(* IEC 61131-3 sources: rusty/tests/lit/single/arithmetic, 10 files *)

(* ---- addition.st ---- *)
// RUN: %COMPILE %s && %RUN | %CHECK %s
// CHECK: 10
FUNCTION main
    VAR
        x : DINT;
        y : DINT;
    END_VAR

    x := 5;
    y := 5;
    printf('%d$N', x + y);
END_FUNCTION

(* ---- integer_overflow.st ---- *)
// RUN: %COMPILE %s && %RUN | %CHECK %s
FUNCTION main
    VAR
        var_sint    : SINT;
        var_int     : INT;
        var_dint    : DINT;
        var_lint    : LINT;

        var_usint   : USINT;
        var_uint    : UINT;
        var_udint   : UDINT;
        var_ulint   : ULINT;
    END_VAR

    // Set max values
    // 8-bit [(2^7)-1]/[(2^8)-1]
    var_sint := 127;                    // Min: -128
    var_usint := 255;                   // Min: 0

    // 16-bit [(2^15)-1]/[(2^16)-1]
    var_int := 32767;                   // Min: -32768
    var_uint := 65535;                  // Min: 0

    // 32-bit [(2^31)-1]/[(2^31)-1]
    var_dint := 2147483647;             // Min: -2147483648
    var_udint := 4294967295;            // Min: 0

    // 64-bit [(2^63)-1]/[(2^64)-1]
    var_lint := 9223372036854775807;    // Min: -9223372036854775808
    var_ulint := 18446744073709551615;  // Min: 0

    // Print and check values
    printf('%d$N', var_sint);       // CHECK: 127
    printf('%d$N', var_int);        // CHECK-NEXT: 32767
    printf('%d$N', var_dint);       // CHECK-NEXT: 2147483647
    printf('%lld$N', var_lint);     // CHECK-NEXT: 9223372036854775807

    printf('%u$N', var_usint);      // CHECK-NEXT: 255
    printf('%u$N', var_uint);       // CHECK-NEXT: 65535
    printf('%u$N', var_udint);      // CHECK-NEXT: 4294967295
    printf('%llu$N', var_ulint);    // CHECK-NEXT: 18446744073709551615

    // Print overflow values
    var_sint := var_sint + 1;
    var_int := var_int + 1;
    var_dint := var_dint + 1;
    var_lint := var_lint + 1;

    var_usint := var_usint + 1;
    var_uint := var_uint + 1;
    var_udint := var_udint + 1;
    var_ulint := var_ulint + 1;

    printf('%d$N', var_sint);       // CHECK: -128
    printf('%d$N', var_int);        // CHECK-NEXT: -32768
    printf('%d$N', var_dint);       // CHECK-NEXT: -2147483648
    printf('%lld$N', var_lint);     // CHECK-NEXT: -9223372036854775808

    printf('%u$N', var_usint);      // CHECK-NEXT: 0
    printf('%u$N', var_uint);       // CHECK-NEXT: 0
    printf('%u$N', var_udint);      // CHECK-NEXT: 0
    printf('%llu$N', var_ulint);    // CHECK-NEXT: 0

END_FUNCTION

(* ---- integer_overflow_with_real_cast.st ---- *)
// RUN: %COMPILE %s && %RUN | %CHECK %s
FUNCTION main
    VAR
        var_int     : INT;
    END_VAR

    printf('%d$N', var_int); // CHECK: 0

    // Cast the REAL value to INT
    var_int := REAL_TO_INT(70_000.4);

    printf('%d$N', var_int); // CHECK: 32767

END_FUNCTION

(* ---- replaced_expression_result_cast.st ---- *)
// RUN: %COMPILE %s && %RUN | %CHECK %s
// The result of a builtin or an operator the compiler carries out through a function call is
// converted to the type of the variable it is assigned to

FUNCTION main
    VAR
        t : TIME := T#10s;
        lt : LTIME := LTIME#10s;
        tod : TOD := TOD#23:59:50;
        n : DINT := 7;
        m : DINT := 3;
        i : INT;
        r : REAL := 2.5;
        x : LREAL;
    END_VAR

    x := t * 1.5;
    printf('%.1f$N', x);                                                            // CHECK: 15000.0
    r := t / 4.0;
    x := r;
    printf('%.1f$N', x);                                                            // CHECK: 2500.0
    x := lt + lt;
    printf('%.1f$N', x);                                                            // CHECK: 20000000000.0

    x := MUL(t, 1.5);
    printf('%.1f$N', x);                                                            // CHECK: 15000.0
    x := ADD(n, m);
    printf('%.1f$N', x);                                                            // CHECK: 10.0
    r := 2.5;
    n := ADD(n, r);
    printf('%d$N', n);                                                              // CHECK: 9
    i := SUB(t, T#4s);
    printf('%d$N', i);                                                              // CHECK: 6000

    tod := (tod + T#20s);
    printf('%s$N', REF(TOD_TO_STRING(tod)));                                        // CHECK: TOD#00:00:10

END_FUNCTION

(* ---- sqrt.st ---- *)
// RUN: %COMPILE %s && %RUN | %CHECK %s
// CHECK: 2
FUNCTION main
    VAR
        res : LREAL;
    END_VAR
    printf('%d$N', REAL_TO_DINT(SQRT(4.0)));
END_FUNCTION

(* ---- unsigned_division_by_literal.st ---- *)
// RUN: %COMPILE %s && %RUN | %CHECK %s
//
// A division of an unsigned operand of 32 or 64 bits by an integer literal is unsigned, like a
// division by a variable of the same type, also when the operand has the highest bit set.

FUNCTION main
    VAR
        udint_value : UDINT := 4_000_000_000;
        two : UDINT := 2;
        dword_value : DWORD := 16#FFFF_FFFF;
        ulint_value : ULINT := 18_446_744_073_709_551_615;
        lword_value : LWORD := 16#FFFF_FFFF_FFFF_FFFF;
    END_VAR
    printf('udint / two: %u$N', udint_value / two);
    printf('udint / 2: %u$N', udint_value / 2);
    printf('dword / 2: %u$N', dword_value / 2);
    printf('ulint / 2: %llu$N', ulint_value / 2);
    printf('lword / 2: %llu$N', lword_value / 2);
    // CHECK:      udint / two: 2000000000
    // CHECK-NEXT: udint / 2: 2000000000
    // CHECK-NEXT: dword / 2: 2147483647
    // CHECK-NEXT: ulint / 2: 9223372036854775807
    // CHECK-NEXT: lword / 2: 9223372036854775807
END_FUNCTION

(* ---- unsigned_division_by_negative_literal.st ---- *)
// RUN: %COMPILE %s && %RUN | %CHECK %s
//
// A negative integer literal does not fit into an unsigned type, so a division or MOD of a UDINT by
// it still runs in DINT and gives a signed result.

FUNCTION main
    VAR
        value : UDINT := 10;
    END_VAR
    printf('value / -2: %d$N', value / -2);
    printf('value MOD -3: %d$N', value MOD -3);
    // CHECK:      value / -2: -5
    // CHECK-NEXT: value MOD -3: 1
END_FUNCTION

(* ---- unsigned_literal_dividend.st ---- *)
// RUN: %COMPILE %s && %RUN | %CHECK %s
//
// An integer literal as the left operand of a division or MOD takes the type of an unsigned divisor of
// 32 bits, so a divisor with the highest bit set is not read as a negative number. As a DINT,
// 16#FFFF_FFFF would be -1, and the results would be -100 and 0.

FUNCTION main
    VAR
        divisor : UDINT := 16#FFFF_FFFF;
    END_VAR
    printf('100 / divisor: %u$N', 100 / divisor);
    printf('100 MOD divisor: %u$N', 100 MOD divisor);
    // CHECK:      100 / divisor: 0
    // CHECK-NEXT: 100 MOD divisor: 100
END_FUNCTION

(* ---- unsigned_modulo_by_literal.st ---- *)
// RUN: %COMPILE %s && %RUN | %CHECK %s
//
// MOD of an unsigned operand of 32 or 64 bits and an integer literal is unsigned, like MOD with a
// variable of the same type, also when the operand has the highest bit set.

FUNCTION main
    VAR
        udint_value : UDINT := 4_000_000_000;
        seven : UDINT := 7;
        dword_value : DWORD := 16#FFFF_FFFF;
        ulint_value : ULINT := 18_446_744_073_709_551_615;
        lword_value : LWORD := 16#FFFF_FFFF_FFFF_FFFF;
    END_VAR
    printf('udint MOD seven: %u$N', udint_value MOD seven);
    printf('udint MOD 7: %u$N', udint_value MOD 7);
    printf('dword MOD 3: %u$N', dword_value MOD 3);
    printf('ulint MOD 10: %llu$N', ulint_value MOD 10);
    printf('lword MOD 10: %llu$N', lword_value MOD 10);
    // CHECK:      udint MOD seven: 3
    // CHECK-NEXT: udint MOD 7: 3
    // CHECK-NEXT: dword MOD 3: 0
    // CHECK-NEXT: ulint MOD 10: 5
    // CHECK-NEXT: lword MOD 10: 5
END_FUNCTION

(* ---- unsigned_subtraction_with_literal.st ---- *)
// RUN: %COMPILE %s && %RUN | %CHECK %s
//
// Addition, subtraction and multiplication of a UDINT and an integer literal still run in DINT, so a
// subtraction below zero gives a negative result instead of wrapping around.

FUNCTION main
    VAR
        value : UDINT := 5;
        wide : LINT;
    END_VAR
    wide := value - 10;
    printf('value - 10: %lld$N', wide);
    printf('value - 10 < 0: %d$N', value - 10 < 0);
    // CHECK:      value - 10: -5
    // CHECK-NEXT: value - 10 < 0: 1
END_FUNCTION
